(* IEC 61131-3 sources: PLC-Static-Analysis/editors/vscode/test/fixtures/project, 2 files *)

(* ---- FB_Pump.st ---- *)
// Pump with a run command.
FUNCTION_BLOCK FB_Pump
VAR_INPUT
    bRun : BOOL; // run command from MAIN
END_VAR
VAR_OUTPUT
    bRunning : BOOL;
END_VAR
bRunning := bRun;
END_FUNCTION_BLOCK

(* ---- MAIN.st ---- *)
PROGRAM MAIN
VAR
    fbPump : FB_Pump;
    rLevel : REAL;
    bAlarm : BOOL;
END_VAR
fbPump(bRun := TRUE);
bAlarm := rLevel = 2.5;
END_PROGRAM
